(* Logix 5000 project; controller TFF vendor 1 type 14 code 107 rev 34.11; software revision 34.03; part 17 of 36 *)
(* tags used below, declared in another part *)
   ControlLoop : ControlLoop[20];   // Control Loop Array
   ControlLoop_PCV001 : ALIAS FOR ControlLoop[3];   // PCV001 Control Loop
   ControlLoop_PCV001_5ms : ALIAS FOR ControlLoop[4];   // PCV001 Control Loop
   ControlLoop_PCV001Alarm : ALIAS FOR AlarmDeviation[3];   // PCV001 Control Loop Deviation Alarm
   ControlLoop_PCV101 : ALIAS FOR ControlLoop[5];   // PCV101 Control Loop
   ControlLoop_PCV101_5ms : ALIAS FOR ControlLoop[6];   // PCV101 Control Loop
   ControlLoop_PCV101_RAMP_OUT : REAL;   // Ramp Output
   PCV001 : ALIAS FOR AnalogPoint[3];   // Retentate Pressure Control Valve Position
   PCV001_AO : ALIAS FOR AnalogOutput[0];   // Retentate Pressure Control Valve Setpoint
   PCV001_Control : PCV_Control;   // PCV001 Control UDT
   PCV001_CVTune : CVTune;
   PCV001_PID : PCV;   // PCV001 PID Management
   PCV101 : ALIAS FOR AnalogPoint[4];   // Filtrate Pressure Control Valve Position
   PCV101_AO : ALIAS FOR AnalogOutput[1];   // FiltratePressure Control Valve Setpoint
   PCV101_Control : PCV_Control;   // PCV101 Control UDT
   PCV101_CVTune : CVTune;
   PCV101_PID : PCV;   // PCV101 PID Management
   Rack_Murr_Node1_TF2S : IO_Station;   // Status of Node 1 TF2S
   Rack_Murr_Node1_TF3S : IO_Station;   // Status of Node 1 TF3S
   RawAnalogInputArray : INT[50];   // Array of analog input raw
   SysControl : SysControl;   // General system status and command
   ThisSystem : SystemType;
   TMP : ALIAS FOR AnalogPoint[41];   // Trans-membrane Pressure
   Valve : Valve[100];   // Valve Array
(* MainProgram5ms, continued *)

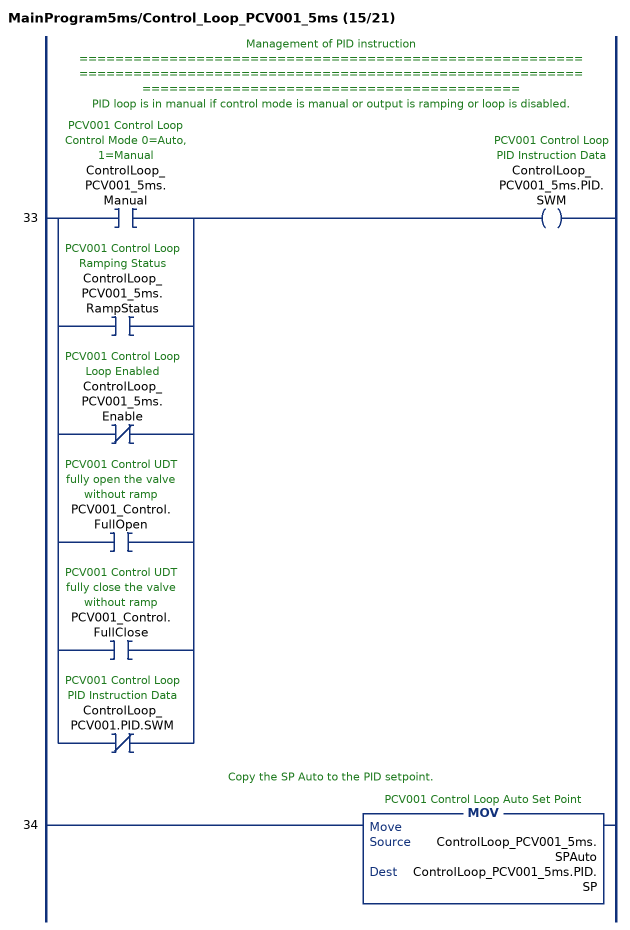
   [picture p67: MainProgram5ms/Control_Loop_PCV001_5ms rungs 33-34]
   // Management of PID instruction
   // ==========================================================================================================================================================
   // PID loop is in manual if control mode is manual or output is ramping or loop is disabled.
   33: [XIC(ControlLoop_PCV001_5ms.Manual) ,XIC(ControlLoop_PCV001_5ms.RampStatus) ,XIO(ControlLoop_PCV001_5ms.Enable) ,[[XIC(PCV001_Control.FullOpen) ,XIC(PCV001_Control.FullClose) ] ,XIO(ControlLoop_PCV001.PID.SWM) ] ]OTE(ControlLoop_PCV001_5ms.PID.SWM);
   // Copy the SP Auto to the PID setpoint.
   34: MOV(ControlLoop_PCV001_5ms.SPAuto,ControlLoop_PCV001_5ms.PID.SP);
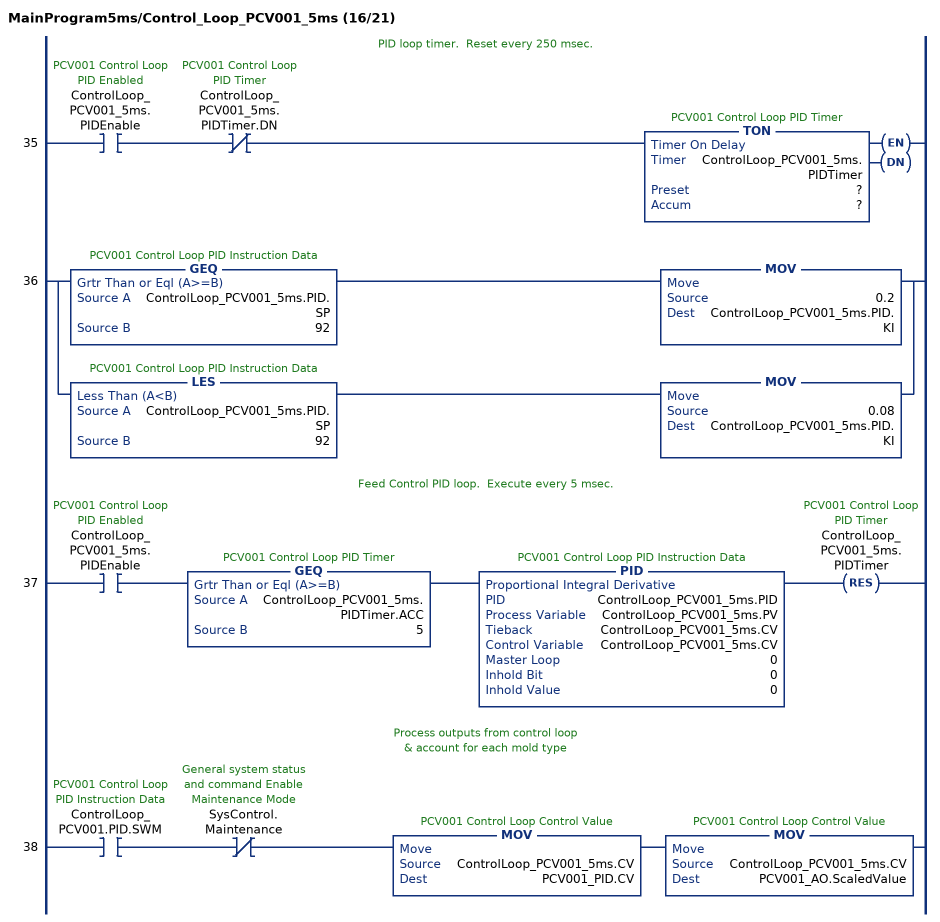
   // PID loop timer.  Reset every 250 msec.
   35: XIC(ControlLoop_PCV001_5ms.PIDEnable)XIO(ControlLoop_PCV001_5ms.PIDTimer.DN)TON(ControlLoop_PCV001_5ms.PIDTimer,?,?);
   36: [GEQ(ControlLoop_PCV001_5ms.PID.SP,92) MOV(0.2,ControlLoop_PCV001_5ms.PID.KI) ,LES(ControlLoop_PCV001_5ms.PID.SP,92) MOV(0.08,ControlLoop_PCV001_5ms.PID.KI) ];
   // Feed Control PID loop.  Execute every 5 msec.
   37: XIC(ControlLoop_PCV001_5ms.PIDEnable)GEQ(ControlLoop_PCV001_5ms.PIDTimer.ACC,5)PID(ControlLoop_PCV001_5ms.PID,ControlLoop_PCV001_5ms.PV,ControlLoop_PCV001_5ms.CV,ControlLoop_PCV001_5ms.CV,0,0,0)RES(ControlLoop_PCV001_5ms.PIDTimer);
   // Process outputs from control loop
   // & account for each mold type
   38: XIC(ControlLoop_PCV001.PID.SWM)XIO(SysControl.Maintenance)MOV(ControlLoop_PCV001_5ms.CV,PCV001_PID.CV)MOV(ControlLoop_PCV001_5ms.CV,PCV001_AO.ScaledValue);
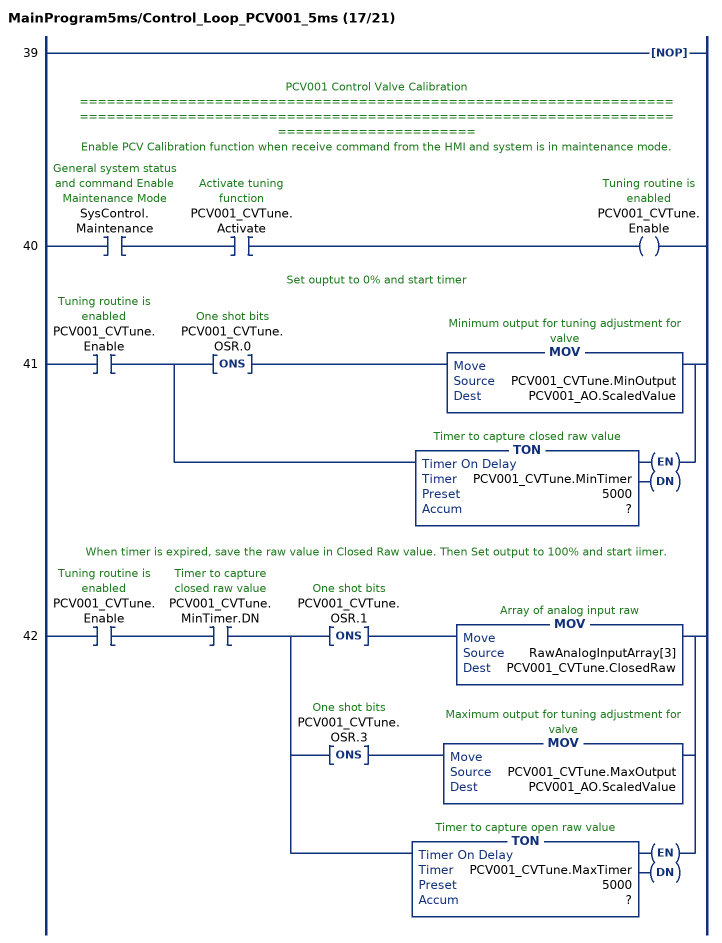
   39: NOP();
   // PCV001 Control Valve Calibration
   // ==========================================================================================================================================================
   // Enable PCV Calibration function when receive command from the HMI and system is in maintenance mode.
   40: XIC(SysControl.Maintenance)XIC(PCV001_CVTune.Activate)OTE(PCV001_CVTune.Enable);
   // Set ouptut to 0% and start timer
   41: XIC(PCV001_CVTune.Enable)[ONS(PCV001_CVTune.OSR.0) MOV(PCV001_CVTune.MinOutput,PCV001_AO.ScaledValue) ,TON(PCV001_CVTune.MinTimer,?,?) ];
   // When timer is expired, save the raw value in Closed Raw value. Then Set output to 100% and start iimer.
   42: XIC(PCV001_CVTune.Enable)XIC(PCV001_CVTune.MinTimer.DN)[ONS(PCV001_CVTune.OSR.1) MOV(RawAnalogInputArray[3],PCV001_CVTune.ClosedRaw) ,ONS(PCV001_CVTune.OSR.3) MOV(PCV001_CVTune.MaxOutput,PCV001_AO.ScaledValue) ,TON(PCV001_CVTune.MaxTimer,?,?) ];
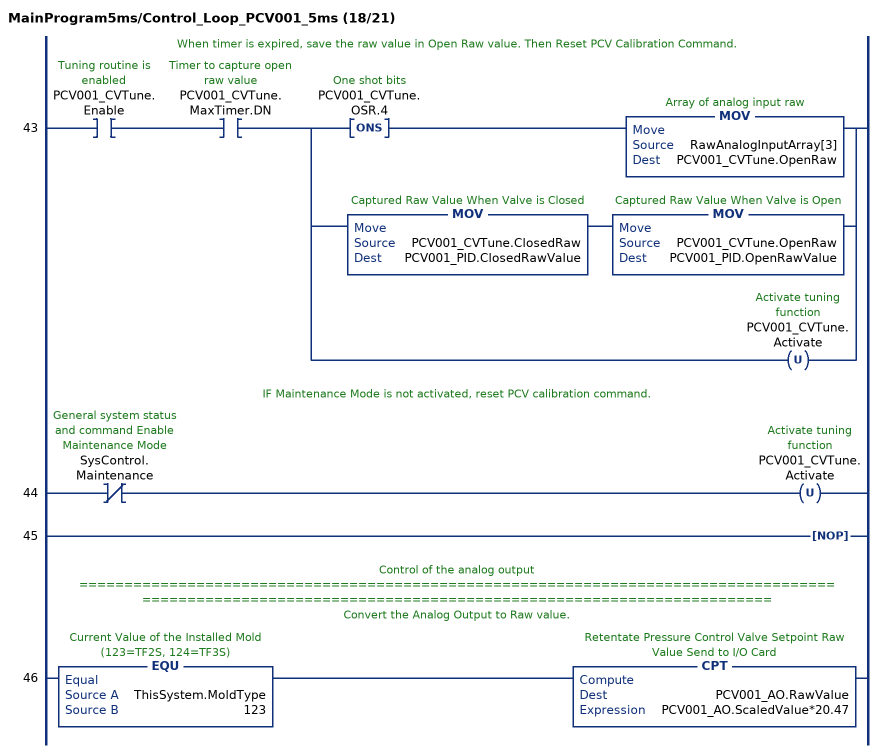
   // When timer is expired, save the raw value in Open Raw value. Then Reset PCV Calibration Command.
   43: XIC(PCV001_CVTune.Enable)XIC(PCV001_CVTune.MaxTimer.DN)[ONS(PCV001_CVTune.OSR.4) MOV(RawAnalogInputArray[3],PCV001_CVTune.OpenRaw) ,MOV(PCV001_CVTune.ClosedRaw,PCV001_PID.ClosedRawValue) MOV(PCV001_CVTune.OpenRaw,PCV001_PID.OpenRawValue) ,OTU(PCV001_CVTune.Activate) ];
   // IF Maintenance Mode is not activated, reset PCV calibration command.
   44: XIO(SysControl.Maintenance)OTU(PCV001_CVTune.Activate);
   45: NOP();
   // Control of the analog output
   // ==========================================================================================================================================================
   // Convert the Analog Output to Raw value.
   46: EQU(ThisSystem.MoldType,123)CPT(PCV001_AO.RawValue,PCV001_AO.ScaledValue*20.47);
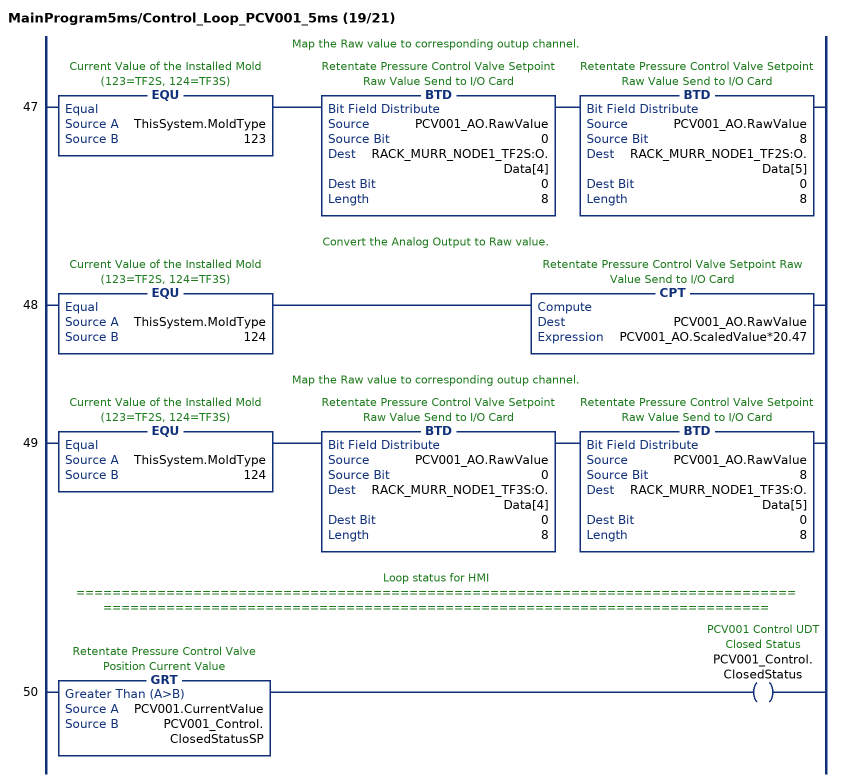
   // Map the Raw value to corresponding outup channel.
   47: EQU(ThisSystem.MoldType,123)BTD(PCV001_AO.RawValue,0,RACK_MURR_NODE1_TF2S:O.Data[4],0,8)BTD(PCV001_AO.RawValue,8,RACK_MURR_NODE1_TF2S:O.Data[5],0,8);
   // Convert the Analog Output to Raw value.
   48: EQU(ThisSystem.MoldType,124)CPT(PCV001_AO.RawValue,PCV001_AO.ScaledValue*20.47);
   // Map the Raw value to corresponding outup channel.
   49: EQU(ThisSystem.MoldType,124)BTD(PCV001_AO.RawValue,0,RACK_MURR_NODE1_TF3S:O.Data[4],0,8)BTD(PCV001_AO.RawValue,8,RACK_MURR_NODE1_TF3S:O.Data[5],0,8);
   // Loop status for HMI
   // ==========================================================================================================================================================
   50: GRT(PCV001.CurrentValue,PCV001_Control.ClosedStatusSP)OTE(PCV001_Control.ClosedStatus);
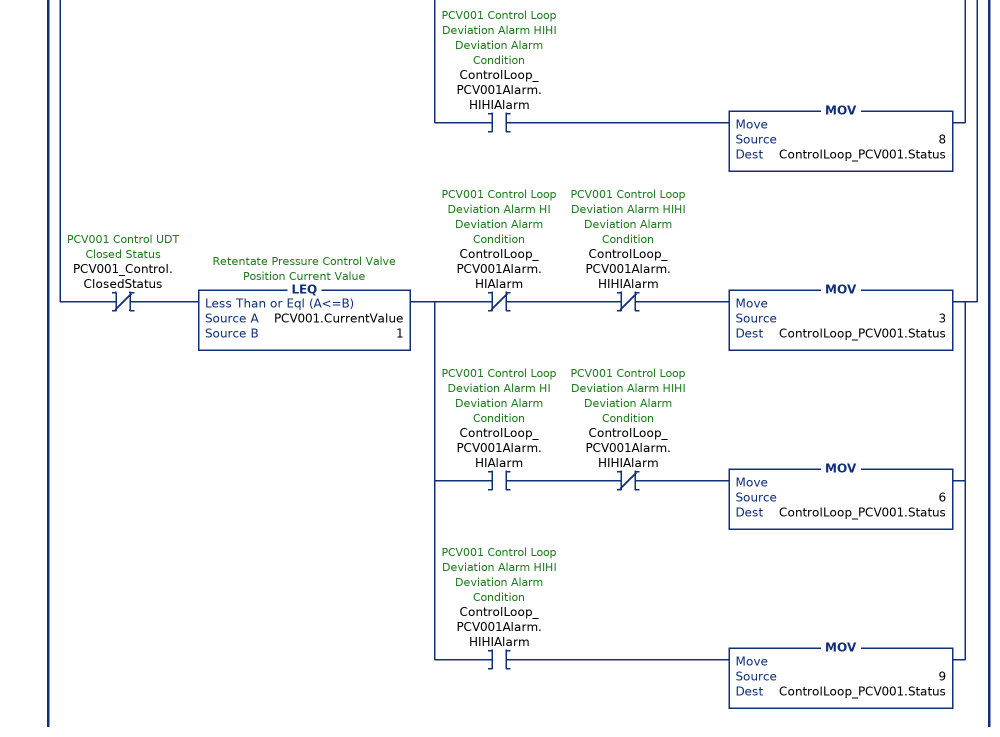
   // ControlLoop Status : 1 = PCV Close
   // ControlLoop Status : 2 = PCV Open
   // ControlLoop Status : 3 = PCV Full Open
   // ControlLoop Status : 4 = PCV Close and Non Critical alam
   // ControlLoop Status : 5 = PCV Open and Non Critical alam
   // ControlLoop Status : 6 = PCV Full Open and Non Critical alam
   // ControlLoop Status : 7 = PCV Close and Critical alam
   // ControlLoop Status : 8 = PCV Open and Critical alam
   // ControlLoop Status : 9 = PCV Full Open and Critical alam
   51: [XIC(PCV001_Control.ClosedStatus) [XIO(ControlLoop_PCV001Alarm.HIAlarm) XIO(ControlLoop_PCV001Alarm.HIHIAlarm) MOV(1,ControlLoop_PCV001.Status) ,XIC(ControlLoop_PCV001Alarm.HIAlarm) XIO(ControlLoop_PCV001Alarm.HIHIAlarm) MOV(4,ControlLoop_PCV001.Status) ,XIC(ControlLoop_PCV001Alarm.HIHIAlarm) MOV(7,ControlLoop_PCV001.Status) ] ,XIO(PCV001_Control.ClosedStatus) GRT(PCV001.CurrentValue,2) [XIO(ControlLoop_PCV001Alarm.HIAlarm) XIO(ControlLoop_PCV001Alarm.HIHIAlarm) MOV(2,ControlLoop_PCV001.Status) ,XIC(ControlLoop_PCV001Alarm.HIAlarm) XIO(ControlLoop_PCV001Alarm.HIHIAlarm) MOV(5,ControlLoop_PCV001.Status) ,XIC(ControlLoop_PCV001Alarm.HIHIAlarm) MOV(8,ControlLoop_PCV001.Status) ] ,XIO(PCV001_Control.ClosedStatus) LEQ(PCV001.CurrentValue,1) [XIO(ControlLoop_PCV001Alarm.HIAlarm) XIO(ControlLoop_PCV001Alarm.HIHIAlarm) MOV(3,ControlLoop_PCV001.Status) ,XIC(ControlLoop_PCV001Alarm.HIAlarm) XIO(ControlLoop_PCV001Alarm.HIHIAlarm) MOV(6,ControlLoop_PCV001.Status) ,XIC(ControlLoop_PCV001Alarm.HIHIAlarm) MOV(9,ControlLoop_PCV001.Status) ] ];
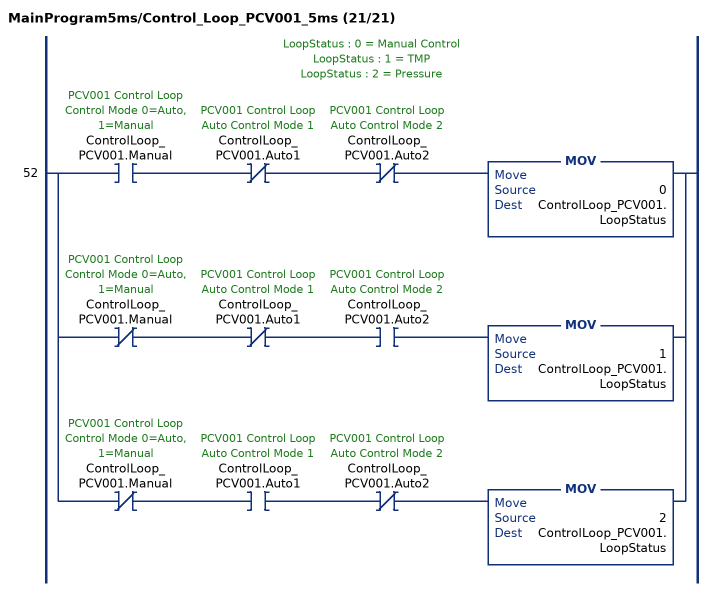
   // LoopStatus : 0 = Manual Control
   //  LoopStatus : 1 = TMP
   //  LoopStatus : 2 = Pressure
   52: [XIC(ControlLoop_PCV001.Manual) XIO(ControlLoop_PCV001.Auto1) XIO(ControlLoop_PCV001.Auto2) MOV(0,ControlLoop_PCV001.LoopStatus) ,XIO(ControlLoop_PCV001.Manual) XIO(ControlLoop_PCV001.Auto1) XIC(ControlLoop_PCV001.Auto2) MOV(1,ControlLoop_PCV001.LoopStatus) ,XIO(ControlLoop_PCV001.Manual) XIC(ControlLoop_PCV001.Auto1) XIO(ControlLoop_PCV001.Auto2) MOV(2,ControlLoop_PCV001.LoopStatus) ];
END_ROUTINE

ROUTINE Control_Loop_PCV101_5ms   (* ladder *)
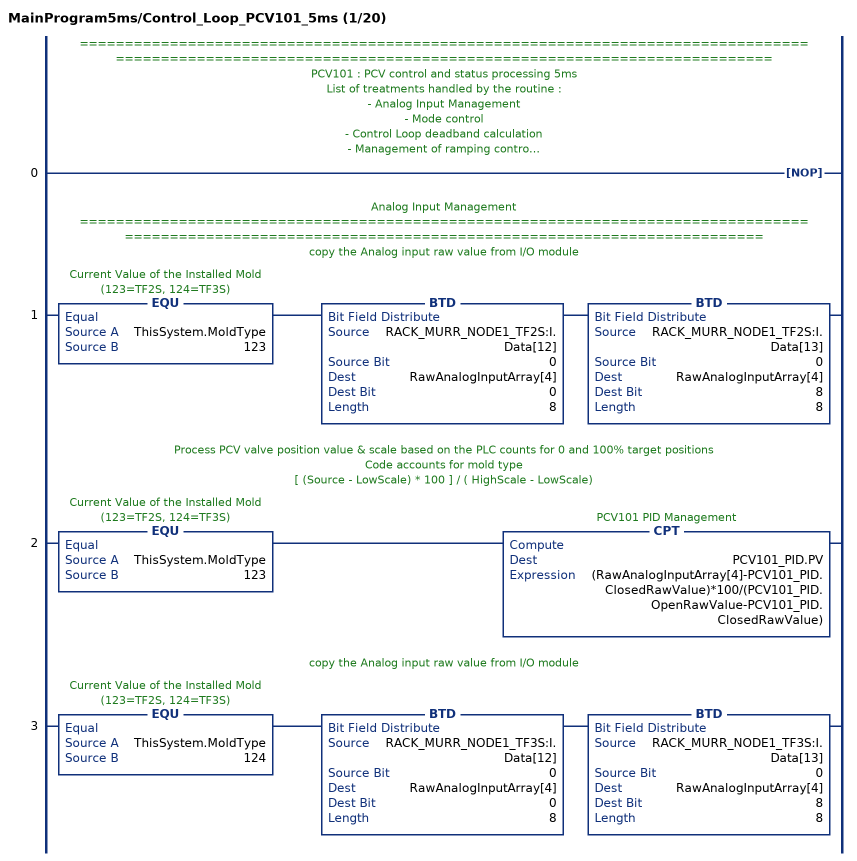
   // ==========================================================================================================================================================
   //                                                  PCV101 : PCV control and status processing 5ms
   //                                                     List of treatments handled by the routine :
   //                                                           - Analog Input Management
   //                                                          - Mode control
   //                                                          - Control Loop deadband calculation
   //                                                          - Management of ramping control
   //                                                          - Management of PID instruction
   //                                                          - PCV101 Control Valve Calibration
   //                                                          - Control of the analog output
   //                                                          - Loop status for HMI
   //                                                     -----------------------------------------------------------------------------------------------------------------------------------------------------
   //                                                     History
   //                                                          2019-AUG-13 - Actemium - B. Roch - Initial version for Candidate Release 3.00.00.00.a
   // 		                                2019-SEP-26 - ACTEMIUM - B. Roch - Modifications for Candidate Release 3.00.00.00.c
   // 					- Change compute for Analog Input Managment
   // 				                                                                - Update Ramping up and down conditions
   // ==========================================================================================================================================================
   0: NOP();
   // Analog Input Management
   // ========================================================================================================================================================
   // copy the Analog input raw value from I/O module
   1: EQU(ThisSystem.MoldType,123)BTD(RACK_MURR_NODE1_TF2S:I.Data[12],0,RawAnalogInputArray[4],0,8)BTD(RACK_MURR_NODE1_TF2S:I.Data[13],0,RawAnalogInputArray[4],8,8);
   // Process PCV valve position value & scale based on the PLC counts for 0 and 100% target positions
   // Code accounts for mold type
   // [ (Source - LowScale) * 100 ] / ( HighScale - LowScale)
   2: EQU(ThisSystem.MoldType,123)CPT(PCV101_PID.PV,(RawAnalogInputArray[4]-PCV101_PID.ClosedRawValue)*100/(PCV101_PID.OpenRawValue-PCV101_PID.ClosedRawValue));
   // copy the Analog input raw value from I/O module
   3: EQU(ThisSystem.MoldType,124)BTD(RACK_MURR_NODE1_TF3S:I.Data[12],0,RawAnalogInputArray[4],0,8)BTD(RACK_MURR_NODE1_TF3S:I.Data[13],0,RawAnalogInputArray[4],8,8);
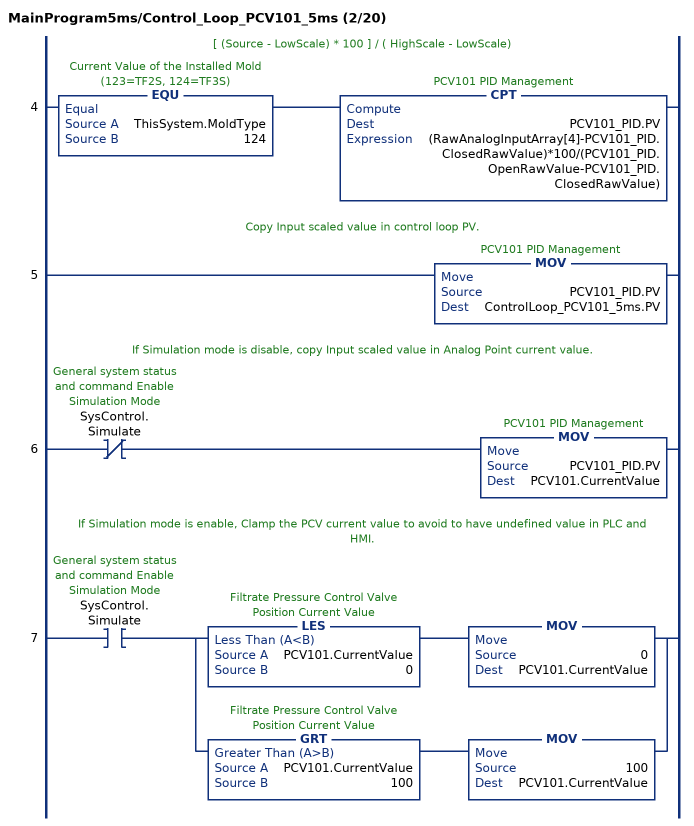
   // [ (Source - LowScale) * 100 ] / ( HighScale - LowScale)
   4: EQU(ThisSystem.MoldType,124)CPT(PCV101_PID.PV,(RawAnalogInputArray[4]-PCV101_PID.ClosedRawValue)*100/(PCV101_PID.OpenRawValue-PCV101_PID.ClosedRawValue));
   // Copy Input scaled value in control loop PV.
   5: MOV(PCV101_PID.PV,ControlLoop_PCV101_5ms.PV);
   // If Simulation mode is disable, copy Input scaled value in Analog Point current value.
   6: XIO(SysControl.Simulate)MOV(PCV101_PID.PV,PCV101.CurrentValue);
   // If Simulation mode is enable, Clamp the PCV current value to avoid to have undefined value in PLC and HMI.
   7: XIC(SysControl.Simulate)[LES(PCV101.CurrentValue,0) MOV(0,PCV101.CurrentValue) ,GRT(PCV101.CurrentValue,100) MOV(100,PCV101.CurrentValue) ];
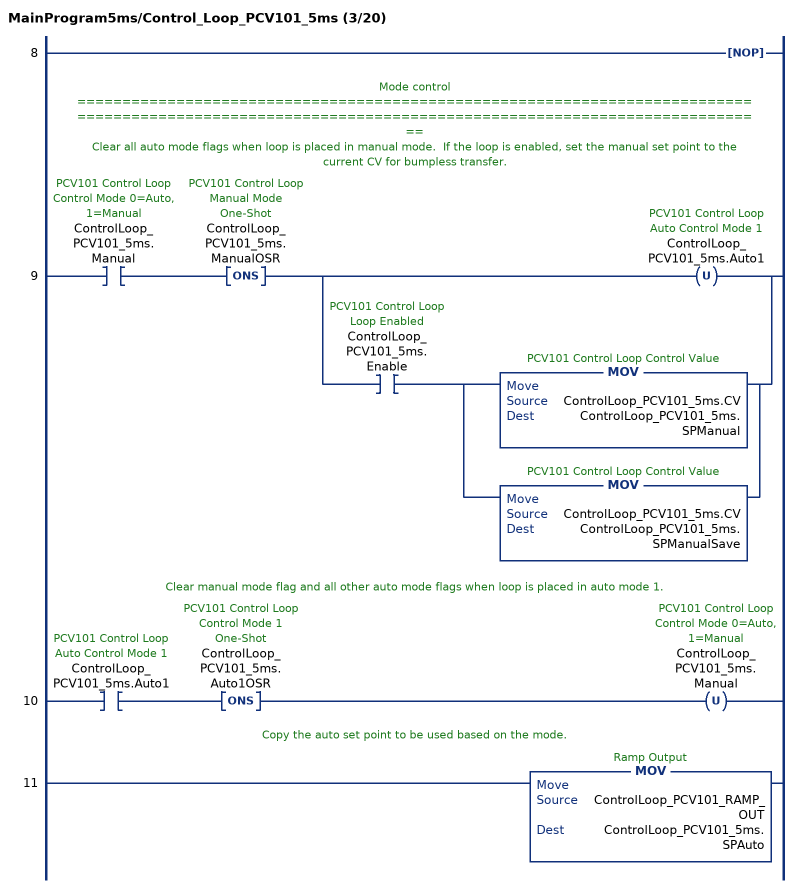
   8: NOP();
   // Mode control
   // ========================================================================================================================================================
   // Clear all auto mode flags when loop is placed in manual mode.  If the loop is enabled, set the manual set point to the current CV for bumpless transfer.
   9: XIC(ControlLoop_PCV101_5ms.Manual)ONS(ControlLoop_PCV101_5ms.ManualOSR)[OTU(ControlLoop_PCV101_5ms.Auto1) ,XIC(ControlLoop_PCV101_5ms.Enable) [MOV(ControlLoop_PCV101_5ms.CV,ControlLoop_PCV101_5ms.SPManual) ,MOV(ControlLoop_PCV101_5ms.CV,ControlLoop_PCV101_5ms.SPManualSave) ] ];
   // Clear manual mode flag and all other auto mode flags when loop is placed in auto mode 1.
   10: XIC(ControlLoop_PCV101_5ms.Auto1)ONS(ControlLoop_PCV101_5ms.Auto1OSR)OTU(ControlLoop_PCV101_5ms.Manual);
   // Copy the auto set point to be used based on the mode.
   11: MOV(ControlLoop_PCV101_RAMP_OUT,ControlLoop_PCV101_5ms.SPAuto);
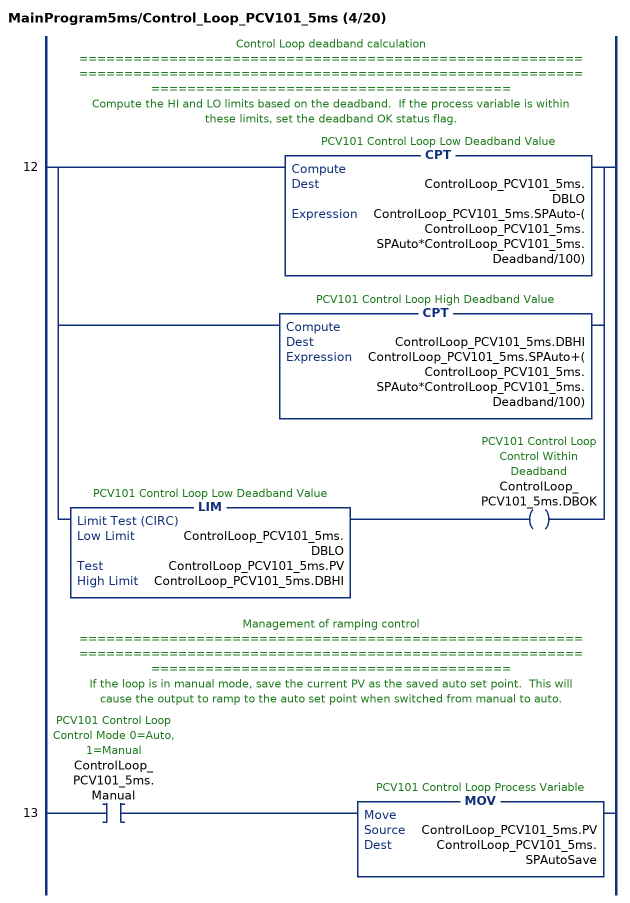
   // Control Loop deadband calculation
   // ========================================================================================================================================================
   // Compute the HI and LO limits based on the deadband.  If the process variable is within these limits, set the deadband OK status flag.
   12: [CPT(ControlLoop_PCV101_5ms.DBLO,ControlLoop_PCV101_5ms.SPAuto-(ControlLoop_PCV101_5ms.SPAuto*ControlLoop_PCV101_5ms.Deadband/100)) ,CPT(ControlLoop_PCV101_5ms.DBHI,ControlLoop_PCV101_5ms.SPAuto+(ControlLoop_PCV101_5ms.SPAuto*ControlLoop_PCV101_5ms.Deadband/100)) ,LIM(ControlLoop_PCV101_5ms.DBLO,ControlLoop_PCV101_5ms.PV,ControlLoop_PCV101_5ms.DBHI) OTE(ControlLoop_PCV101_5ms.DBOK) ];
   // Management of ramping control
   // ========================================================================================================================================================
   // If the loop is in manual mode, save the current PV as the saved auto set point.  This will cause the output to ramp to the auto set point when switched from manual to auto.
   13: XIC(ControlLoop_PCV101_5ms.Manual)MOV(ControlLoop_PCV101_5ms.PV,ControlLoop_PCV101_5ms.SPAutoSave);
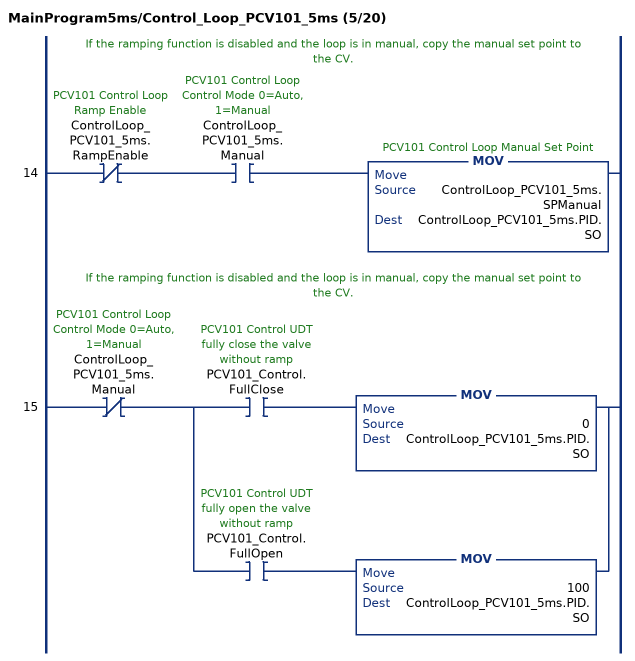
   // If the ramping function is disabled and the loop is in manual, copy the manual set point to the CV.
   14: XIO(ControlLoop_PCV101_5ms.RampEnable)XIC(ControlLoop_PCV101_5ms.Manual)MOV(ControlLoop_PCV101_5ms.SPManual,ControlLoop_PCV101_5ms.PID.SO);
   // If the ramping function is disabled and the loop is in manual, copy the manual set point to the CV.
   15: XIO(ControlLoop_PCV101_5ms.Manual)[XIC(PCV101_Control.FullClose) MOV(0,ControlLoop_PCV101_5ms.PID.SO) ,XIC(PCV101_Control.FullOpen) MOV(100,ControlLoop_PCV101_5ms.PID.SO) ];
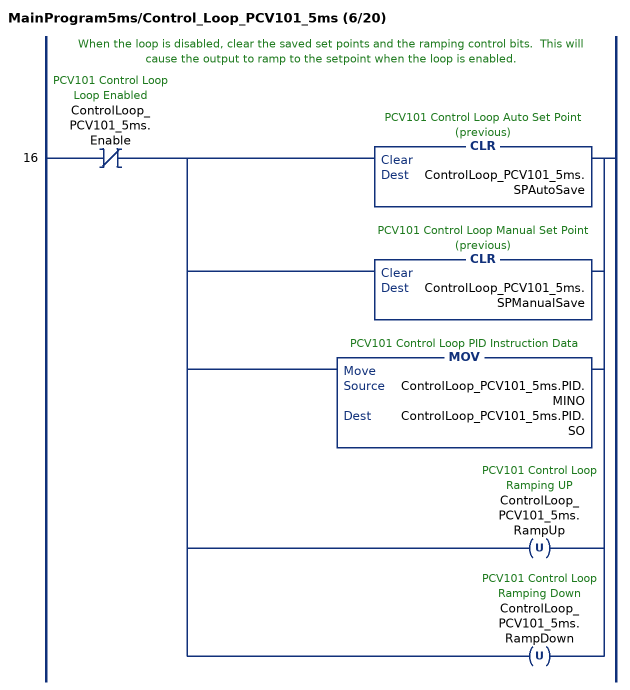
   // When the loop is disabled, clear the saved set points and the ramping control bits.  This will cause the output to ramp to the setpoint when the loop is enabled.
   16: XIO(ControlLoop_PCV101_5ms.Enable)[CLR(ControlLoop_PCV101_5ms.SPAutoSave) ,CLR(ControlLoop_PCV101_5ms.SPManualSave) ,MOV(ControlLoop_PCV101_5ms.PID.MINO,ControlLoop_PCV101_5ms.PID.SO) ,OTU(ControlLoop_PCV101_5ms.RampUp) ,OTU(ControlLoop_PCV101_5ms.RampDown) ];
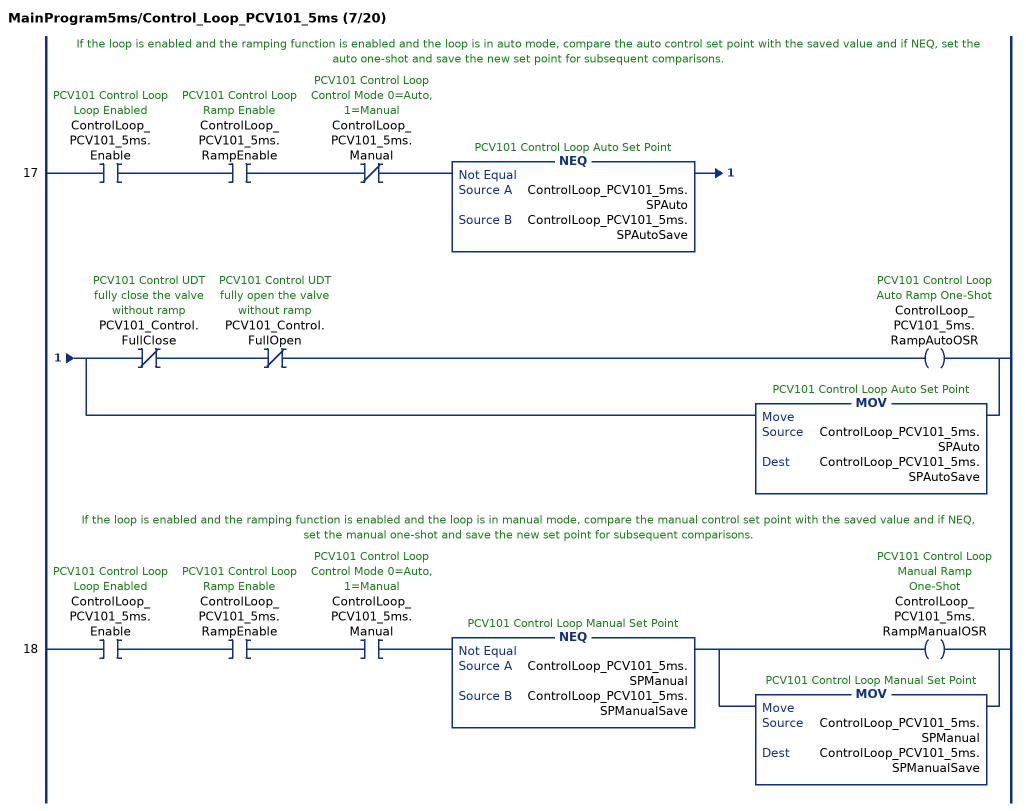
   // If the loop is enabled and the ramping function is enabled and the loop is in auto mode, compare the auto control set point with the saved value and if NEQ, set the auto one-shot and save the new set point for subsequent comparisons.
   17: XIC(ControlLoop_PCV101_5ms.Enable)XIC(ControlLoop_PCV101_5ms.RampEnable)XIO(ControlLoop_PCV101_5ms.Manual)NEQ(ControlLoop_PCV101_5ms.SPAuto,ControlLoop_PCV101_5ms.SPAutoSave)[XIO(PCV101_Control.FullClose) XIO(PCV101_Control.FullOpen) OTE(ControlLoop_PCV101_5ms.RampAutoOSR) ,MOV(ControlLoop_PCV101_5ms.SPAuto,ControlLoop_PCV101_5ms.SPAutoSave) ];
   // If the loop is enabled and the ramping function is enabled and the loop is in manual mode, compare the manual control set point with the saved value and if NEQ, set the manual one-shot and save the new set point for subsequent comparisons.
   18: XIC(ControlLoop_PCV101_5ms.Enable)XIC(ControlLoop_PCV101_5ms.RampEnable)XIC(ControlLoop_PCV101_5ms.Manual)NEQ(ControlLoop_PCV101_5ms.SPManual,ControlLoop_PCV101_5ms.SPManualSave)[OTE(ControlLoop_PCV101_5ms.RampManualOSR) ,MOV(ControlLoop_PCV101_5ms.SPManual,ControlLoop_PCV101_5ms.SPManualSave) ];
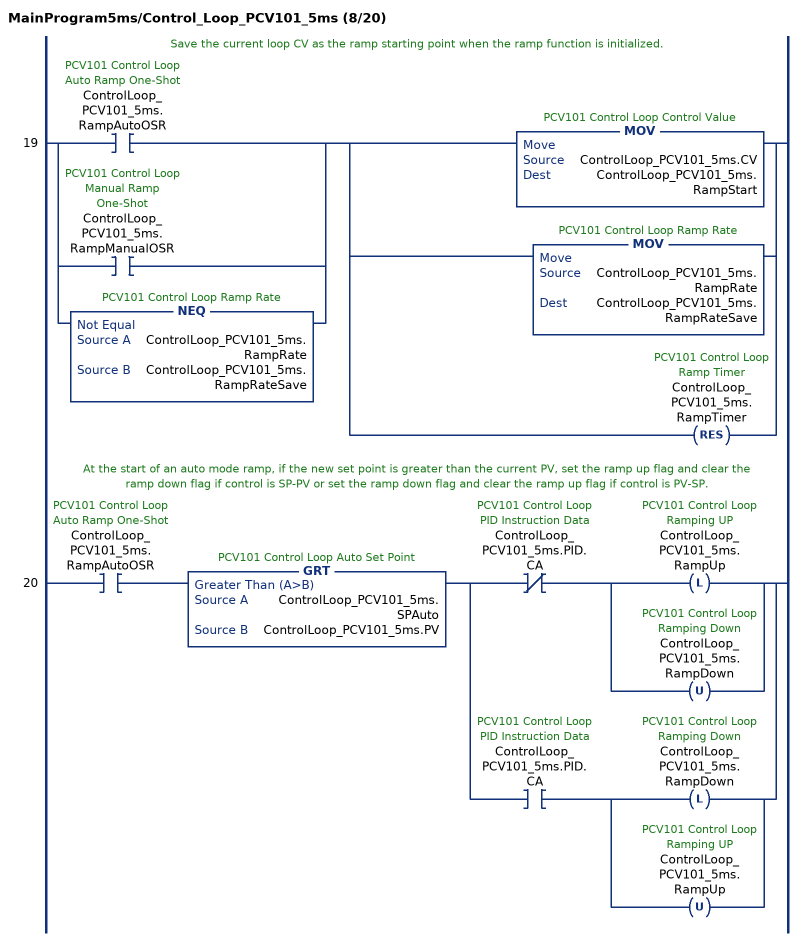
   // Save the current loop CV as the ramp starting point when the ramp function is initialized.
   19: [XIC(ControlLoop_PCV101_5ms.RampAutoOSR) ,XIC(ControlLoop_PCV101_5ms.RampManualOSR) ,NEQ(ControlLoop_PCV101_5ms.RampRate,ControlLoop_PCV101_5ms.RampRateSave) ][MOV(ControlLoop_PCV101_5ms.CV,ControlLoop_PCV101_5ms.RampStart) ,MOV(ControlLoop_PCV101_5ms.RampRate,ControlLoop_PCV101_5ms.RampRateSave) ,RES(ControlLoop_PCV101_5ms.RampTimer) ];
   // At the start of an auto mode ramp, if the new set point is greater than the current PV, set the ramp up flag and clear the ramp down flag if control is SP-PV or set the ramp down flag and clear the ramp up flag if control is PV-SP.
   20: XIC(ControlLoop_PCV101_5ms.RampAutoOSR)GRT(ControlLoop_PCV101_5ms.SPAuto,ControlLoop_PCV101_5ms.PV)[XIO(ControlLoop_PCV101_5ms.PID.CA) [OTL(ControlLoop_PCV101_5ms.RampUp) ,OTU(ControlLoop_PCV101_5ms.RampDown) ] ,XIC(ControlLoop_PCV101_5ms.PID.CA) [OTL(ControlLoop_PCV101_5ms.RampDown) ,OTU(ControlLoop_PCV101_5ms.RampUp) ] ];
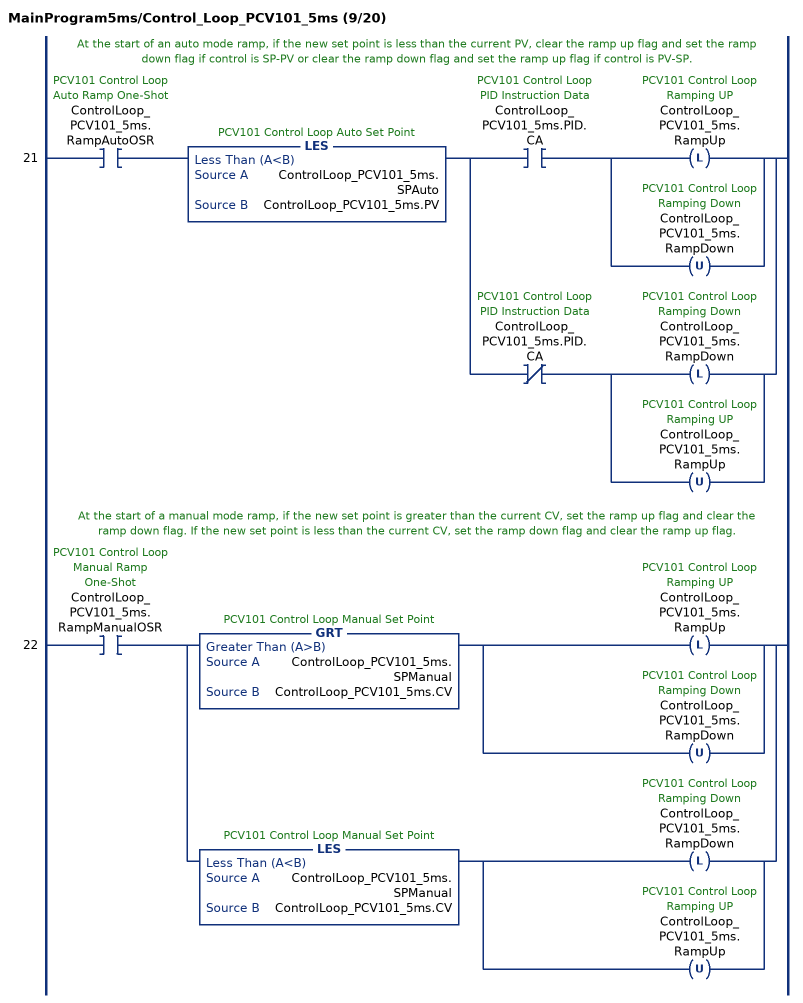
   // At the start of an auto mode ramp, if the new set point is less than the current PV, clear the ramp up flag and set the ramp down flag if control is SP-PV or clear the ramp down flag and set the ramp up flag if control is PV-SP.
   21: XIC(ControlLoop_PCV101_5ms.RampAutoOSR)LES(ControlLoop_PCV101_5ms.SPAuto,ControlLoop_PCV101_5ms.PV)[XIC(ControlLoop_PCV101_5ms.PID.CA) [OTL(ControlLoop_PCV101_5ms.RampUp) ,OTU(ControlLoop_PCV101_5ms.RampDown) ] ,XIO(ControlLoop_PCV101_5ms.PID.CA) [OTL(ControlLoop_PCV101_5ms.RampDown) ,OTU(ControlLoop_PCV101_5ms.RampUp) ] ];
   // At the start of a manual mode ramp, if the new set point is greater than the current CV, set the ramp up flag and clear the ramp down flag. If the new set point is less than the current CV, set the ramp down flag and clear the ramp up flag.
   22: XIC(ControlLoop_PCV101_5ms.RampManualOSR)[GRT(ControlLoop_PCV101_5ms.SPManual,ControlLoop_PCV101_5ms.CV) [OTL(ControlLoop_PCV101_5ms.RampUp) ,OTU(ControlLoop_PCV101_5ms.RampDown) ] ,LES(ControlLoop_PCV101_5ms.SPManual,ControlLoop_PCV101_5ms.CV) [OTL(ControlLoop_PCV101_5ms.RampDown) ,OTU(ControlLoop_PCV101_5ms.RampUp) ] ];
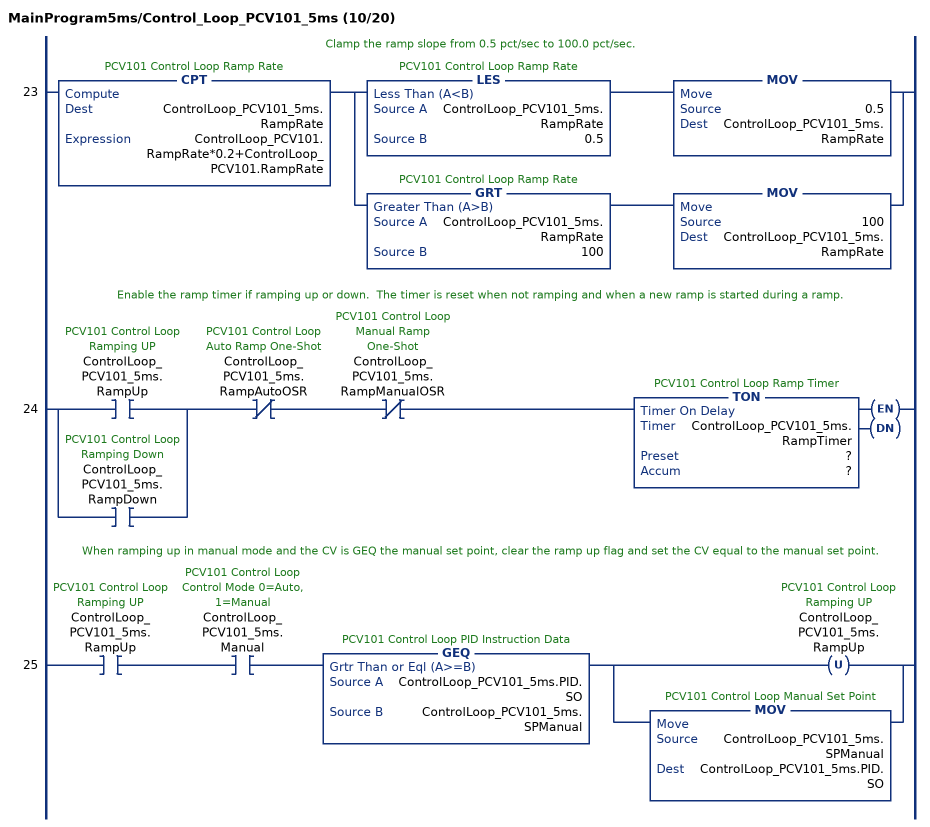
   // Clamp the ramp slope from 0.5 pct/sec to 100.0 pct/sec.
   23: CPT(ControlLoop_PCV101_5ms.RampRate,ControlLoop_PCV101.RampRate*0.2+ControlLoop_PCV101.RampRate)[LES(ControlLoop_PCV101_5ms.RampRate,0.5) MOV(0.5,ControlLoop_PCV101_5ms.RampRate) ,GRT(ControlLoop_PCV101_5ms.RampRate,100) MOV(100,ControlLoop_PCV101_5ms.RampRate) ];
   // Enable the ramp timer if ramping up or down.  The timer is reset when not ramping and when a new ramp is started during a ramp.
   24: [XIC(ControlLoop_PCV101_5ms.RampUp) ,XIC(ControlLoop_PCV101_5ms.RampDown) ]XIO(ControlLoop_PCV101_5ms.RampAutoOSR)XIO(ControlLoop_PCV101_5ms.RampManualOSR)TON(ControlLoop_PCV101_5ms.RampTimer,?,?);
   // When ramping up in manual mode and the CV is GEQ the manual set point, clear the ramp up flag and set the CV equal to the manual set point.
   25: XIC(ControlLoop_PCV101_5ms.RampUp)XIC(ControlLoop_PCV101_5ms.Manual)GEQ(ControlLoop_PCV101_5ms.PID.SO,ControlLoop_PCV101_5ms.SPManual)[OTU(ControlLoop_PCV101_5ms.RampUp) ,MOV(ControlLoop_PCV101_5ms.SPManual,ControlLoop_PCV101_5ms.PID.SO) ];
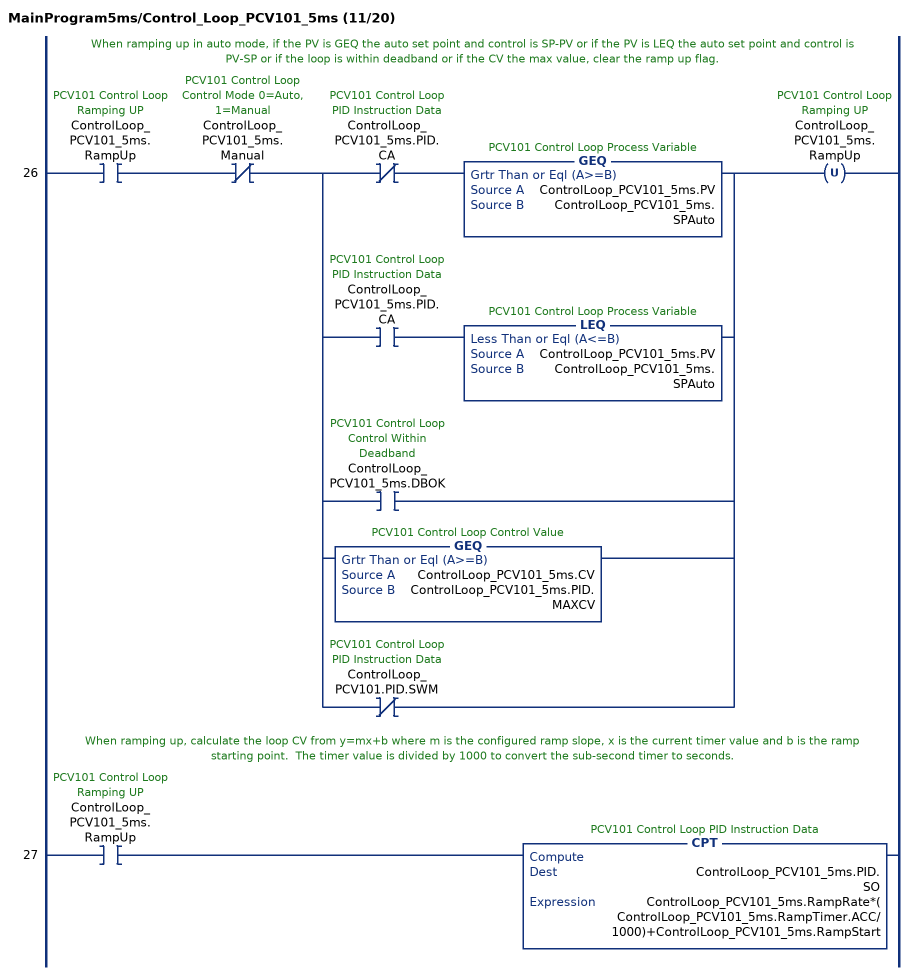
   // When ramping up in auto mode, if the PV is GEQ the auto set point and control is SP-PV or if the PV is LEQ the auto set point and control is PV-SP or if the loop is within deadband or if the CV the max value, clear the ramp up flag.
   26: XIC(ControlLoop_PCV101_5ms.RampUp)XIO(ControlLoop_PCV101_5ms.Manual)[XIO(ControlLoop_PCV101_5ms.PID.CA) GEQ(ControlLoop_PCV101_5ms.PV,ControlLoop_PCV101_5ms.SPAuto) ,XIC(ControlLoop_PCV101_5ms.PID.CA) LEQ(ControlLoop_PCV101_5ms.PV,ControlLoop_PCV101_5ms.SPAuto) ,XIC(ControlLoop_PCV101_5ms.DBOK) ,[GEQ(ControlLoop_PCV101_5ms.CV,ControlLoop_PCV101_5ms.PID.MAXCV) ,XIO(ControlLoop_PCV101.PID.SWM) ] ]OTU(ControlLoop_PCV101_5ms.RampUp);
   // When ramping up, calculate the loop CV from y=mx+b where m is the configured ramp slope, x is the current timer value and b is the ramp starting point.  The timer value is divided by 1000 to convert the sub-second timer to seconds.
   27: XIC(ControlLoop_PCV101_5ms.RampUp)CPT(ControlLoop_PCV101_5ms.PID.SO,ControlLoop_PCV101_5ms.RampRate*(ControlLoop_PCV101_5ms.RampTimer.ACC/1000)+ControlLoop_PCV101_5ms.RampStart);
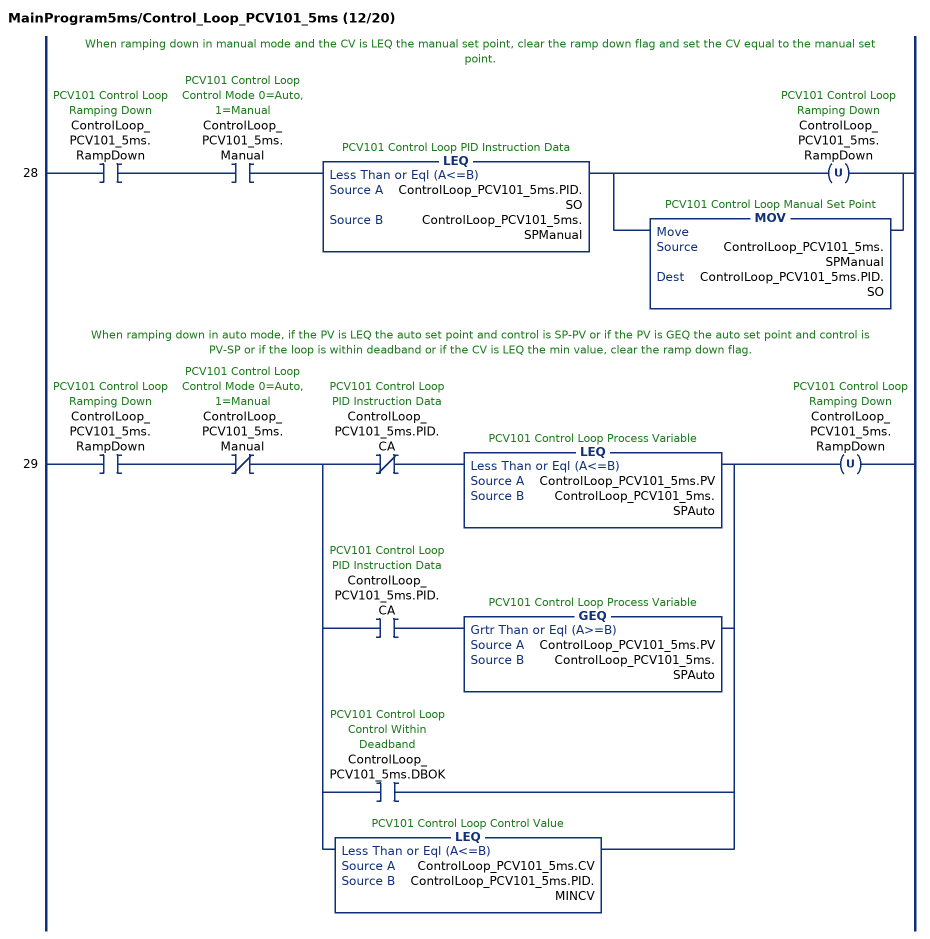
   // When ramping down in manual mode and the CV is LEQ the manual set point, clear the ramp down flag and set the CV equal to the manual set point.
   28: XIC(ControlLoop_PCV101_5ms.RampDown)XIC(ControlLoop_PCV101_5ms.Manual)LEQ(ControlLoop_PCV101_5ms.PID.SO,ControlLoop_PCV101_5ms.SPManual)[OTU(ControlLoop_PCV101_5ms.RampDown) ,MOV(ControlLoop_PCV101_5ms.SPManual,ControlLoop_PCV101_5ms.PID.SO) ];
   // When ramping down in auto mode, if the PV is LEQ the auto set point and control is SP-PV or if the PV is GEQ the auto set point and control is PV-SP or if the loop is within deadband or if the CV is LEQ the min value, clear the ramp down flag.
   29: XIC(ControlLoop_PCV101_5ms.RampDown)XIO(ControlLoop_PCV101_5ms.Manual)[XIO(ControlLoop_PCV101_5ms.PID.CA) LEQ(ControlLoop_PCV101_5ms.PV,ControlLoop_PCV101_5ms.SPAuto) ,XIC(ControlLoop_PCV101_5ms.PID.CA) GEQ(ControlLoop_PCV101_5ms.PV,ControlLoop_PCV101_5ms.SPAuto) ,XIC(ControlLoop_PCV101_5ms.DBOK) ,LEQ(ControlLoop_PCV101_5ms.CV,ControlLoop_PCV101_5ms.PID.MINCV) ]OTU(ControlLoop_PCV101_5ms.RampDown);
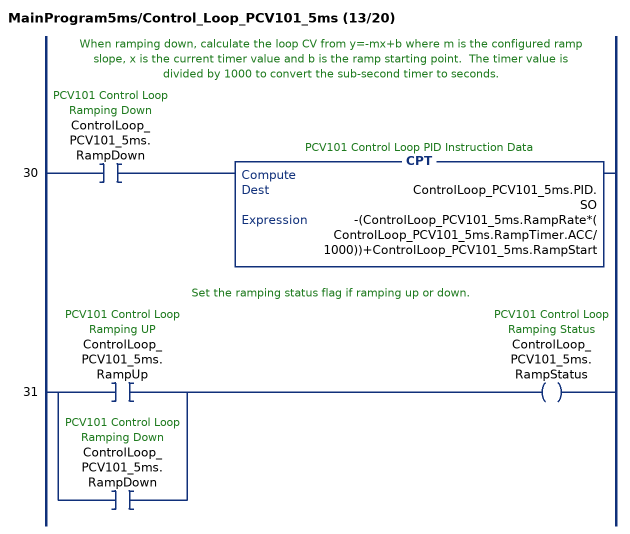
   // When ramping down, calculate the loop CV from y=-mx+b where m is the configured ramp slope, x is the current timer value and b is the ramp starting point.  The timer value is divided by 1000 to convert the sub-second timer to seconds.
   30: XIC(ControlLoop_PCV101_5ms.RampDown)CPT(ControlLoop_PCV101_5ms.PID.SO,-(ControlLoop_PCV101_5ms.RampRate*(ControlLoop_PCV101_5ms.RampTimer.ACC/1000))+ControlLoop_PCV101_5ms.RampStart);
   // Set the ramping status flag if ramping up or down.
   31: [XIC(ControlLoop_PCV101_5ms.RampUp) ,XIC(ControlLoop_PCV101_5ms.RampDown) ]OTE(ControlLoop_PCV101_5ms.RampStatus);
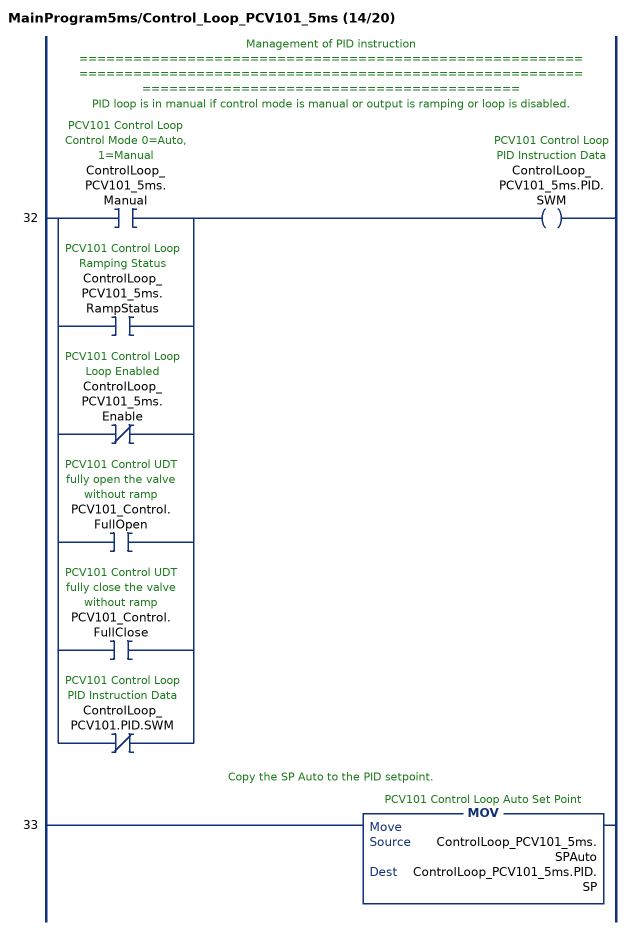
   // Management of PID instruction
   // ==========================================================================================================================================================
   // PID loop is in manual if control mode is manual or output is ramping or loop is disabled.
   32: [XIC(ControlLoop_PCV101_5ms.Manual) ,XIC(ControlLoop_PCV101_5ms.RampStatus) ,XIO(ControlLoop_PCV101_5ms.Enable) ,[[XIC(PCV101_Control.FullOpen) ,XIC(PCV101_Control.FullClose) ] ,XIO(ControlLoop_PCV101.PID.SWM) ] ]OTE(ControlLoop_PCV101_5ms.PID.SWM);
   // Copy the SP Auto to the PID setpoint.
   33: MOV(ControlLoop_PCV101_5ms.SPAuto,ControlLoop_PCV101_5ms.PID.SP);
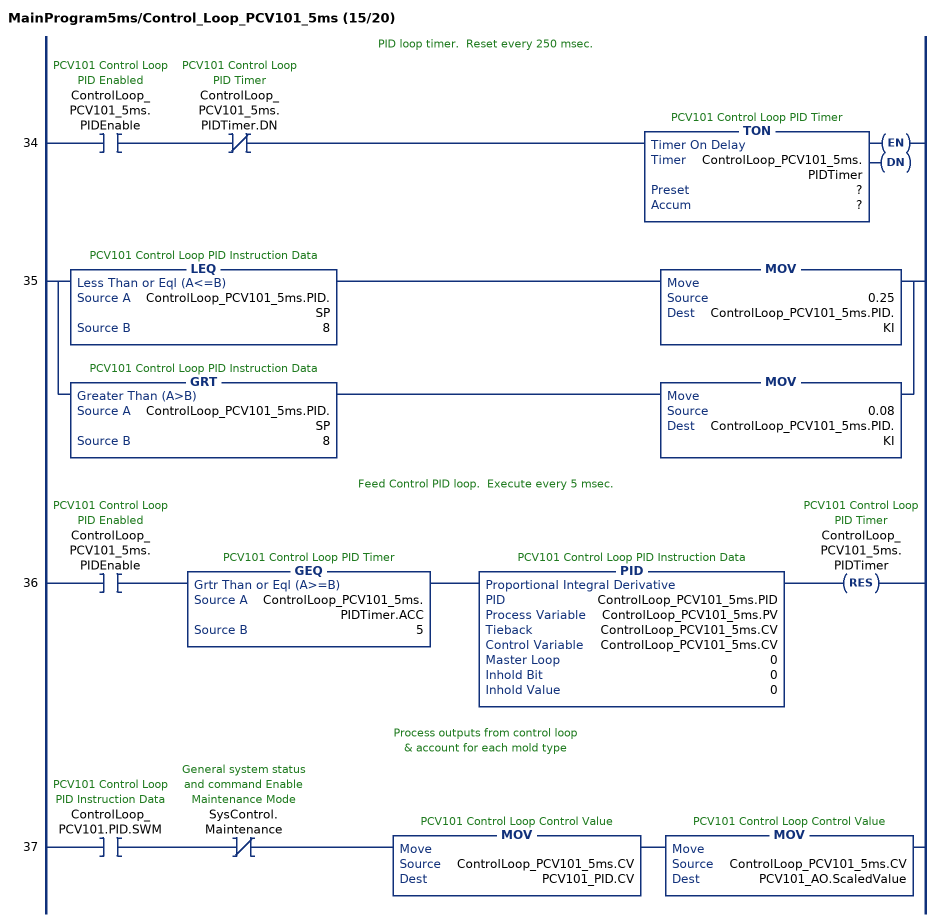
   // PID loop timer.  Reset every 250 msec.
   34: XIC(ControlLoop_PCV101_5ms.PIDEnable)XIO(ControlLoop_PCV101_5ms.PIDTimer.DN)TON(ControlLoop_PCV101_5ms.PIDTimer,?,?);
   35: [LEQ(ControlLoop_PCV101_5ms.PID.SP,8) MOV(0.25,ControlLoop_PCV101_5ms.PID.KI) ,GRT(ControlLoop_PCV101_5ms.PID.SP,8) MOV(0.08,ControlLoop_PCV101_5ms.PID.KI) ];
   // Feed Control PID loop.  Execute every 5 msec.
   36: XIC(ControlLoop_PCV101_5ms.PIDEnable)GEQ(ControlLoop_PCV101_5ms.PIDTimer.ACC,5)PID(ControlLoop_PCV101_5ms.PID,ControlLoop_PCV101_5ms.PV,ControlLoop_PCV101_5ms.CV,ControlLoop_PCV101_5ms.CV,0,0,0)RES(ControlLoop_PCV101_5ms.PIDTimer);
   // Process outputs from control loop
   // & account for each mold type
   37: XIC(ControlLoop_PCV101.PID.SWM)XIO(SysControl.Maintenance)MOV(ControlLoop_PCV101_5ms.CV,PCV101_PID.CV)MOV(ControlLoop_PCV101_5ms.CV,PCV101_AO.ScaledValue);
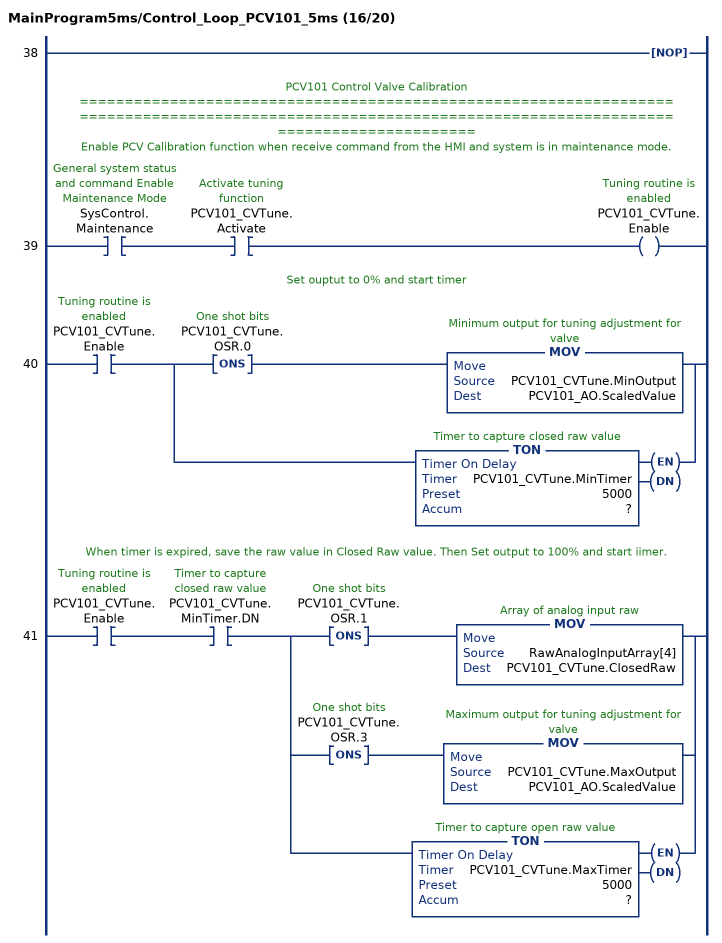
   38: NOP();
   // PCV101 Control Valve Calibration
   // ==========================================================================================================================================================
   // Enable PCV Calibration function when receive command from the HMI and system is in maintenance mode.
   39: XIC(SysControl.Maintenance)XIC(PCV101_CVTune.Activate)OTE(PCV101_CVTune.Enable);
   // Set ouptut to 0% and start timer
   40: XIC(PCV101_CVTune.Enable)[ONS(PCV101_CVTune.OSR.0) MOV(PCV101_CVTune.MinOutput,PCV101_AO.ScaledValue) ,TON(PCV101_CVTune.MinTimer,?,?) ];
   // When timer is expired, save the raw value in Closed Raw value. Then Set output to 100% and start iimer.
   41: XIC(PCV101_CVTune.Enable)XIC(PCV101_CVTune.MinTimer.DN)[ONS(PCV101_CVTune.OSR.1) MOV(RawAnalogInputArray[4],PCV101_CVTune.ClosedRaw) ,ONS(PCV101_CVTune.OSR.3) MOV(PCV101_CVTune.MaxOutput,PCV101_AO.ScaledValue) ,TON(PCV101_CVTune.MaxTimer,?,?) ];
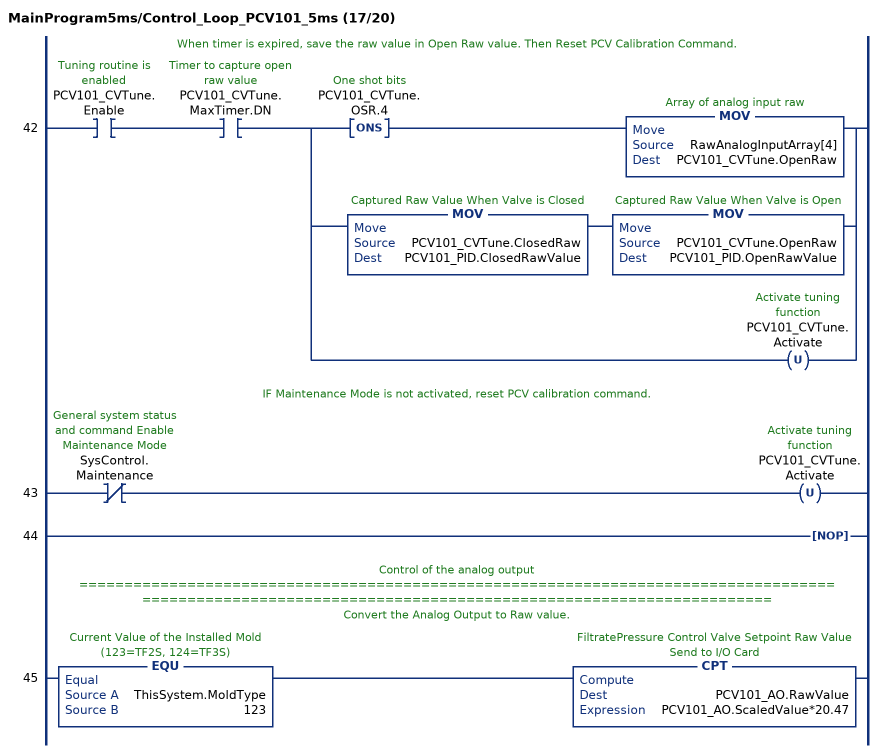
   // When timer is expired, save the raw value in Open Raw value. Then Reset PCV Calibration Command.
   42: XIC(PCV101_CVTune.Enable)XIC(PCV101_CVTune.MaxTimer.DN)[ONS(PCV101_CVTune.OSR.4) MOV(RawAnalogInputArray[4],PCV101_CVTune.OpenRaw) ,MOV(PCV101_CVTune.ClosedRaw,PCV101_PID.ClosedRawValue) MOV(PCV101_CVTune.OpenRaw,PCV101_PID.OpenRawValue) ,OTU(PCV101_CVTune.Activate) ];
   // IF Maintenance Mode is not activated, reset PCV calibration command.
   43: XIO(SysControl.Maintenance)OTU(PCV101_CVTune.Activate);
   44: NOP();
   // Control of the analog output
   // ==========================================================================================================================================================
   // Convert the Analog Output to Raw value.
   45: EQU(ThisSystem.MoldType,123)CPT(PCV101_AO.RawValue,PCV101_AO.ScaledValue*20.47);
